(* IEC 61131-3 sources: s7-to-codesys/src/POUs/Lang/Converted/FB_PumpInterlockLad, 2 files *)

(* ---- FB_PumpInterlockLad.decl.st ---- *)
// Назначение: Блокировки насоса по уровню и давлению (LAD)
//             Блокировки насоса II подъёма по уровню в РЧВ и давлению в коллекторе (LAD).
//             1. xLowLevel := iLevel_cm < iLevelMin_cm.  2. xHighPress := iPressure_kPa > iPressureMax_kPa.
//             3. Если xLowLevel OR xHighPress — установить xAlarmLatch (S).
//             4. Если xAck AND NOT xLowLevel AND NOT xHighPress — сбросить xAlarmLatch (R).
//             5. Обслуживание: при xMaint прыжок вперёд к метке NoAuto (сети 6-7 не выполняются).
//             6. xPumpOn := xAutoReq AND NOT xAlarmLatch.
//             7. По фронту xPumpOn (P_TRIG, бит xRunEdge): iRunCount := iRunCount + 1 (ADD Int); xCountOk := ENO
//             сложения
//             (ENO = 0 при переполнении Int: 32767 + 1).
// Автор:      WTP2 (исходный блок S7); перевод в ST — s7conv 0.1.0
// Версия:     0.1 (исходный блок S7)
// Документ:   docs/CONVERSION_REPORT.md, docs/MAPPING.md
// Источник:   samples/lang/FB_PumpInterlockLad.xml, LAD, SW.Blocks.FB "FB_PumpInterlockLad", пространство имён
//             Interface/v5, FAMILY Drives
// Сгенерировано s7conv: пометки MIGRATION-CHECK и MIGRATION-TODO требуют ручного разбора.
FUNCTION_BLOCK FB_PumpInterlockLad
VAR_INPUT
    xAutoReq : BOOL;  // Запрос автоматики на работу
    iLevel_cm : INT;  // Уровень в РЧВ, см
    iLevelMin_cm : INT := 50;  // Минимальный уровень, см
    iPressure_kPa : INT;  // Давление в коллекторе, кПа
    iPressureMax_kPa : INT := 600;  // Максимальное давление, кПа
    xAck : BOOL;  // Квитирование аварии
    xMaint : BOOL;  // Режим обслуживания
END_VAR
VAR_OUTPUT
    xPumpOn : BOOL;  // Команда насосу
    xLowLevel : BOOL;  // Низкий уровень
    xHighPress : BOOL;  // Высокое давление
    xAlarm : BOOL;  // Авария (защёлка)
    iRunCount : INT;  // Число включений
    xCountOk : BOOL;  // ENO сложения: нет переполнения
    iSetpoint_pct : INT;  // Уставка производительности, %
    xChainOk : BOOL;  // ENO цепочки вызовов
    xRunMem : BOOL;  // Копия бита памяти фронта
END_VAR
VAR
    xAlarmLatch : BOOL;  // Защёлка аварии
    xRunEdge : BOOL;  // Бит памяти фронта xPumpOn
    iStage1 : INT;  // Уставка после первого ограничения
    iStage2 : INT;  // Уставка после второго ограничения
END_VAR
VAR_TEMP
    xNet5_1 : BOOL;  // сеть 5: условие прыжка к NoAuto (UId 21)
    xNet7_1 : BOOL;  // сеть 7: PBox (UId 21)
    xNet7_2 : BOOL;  // сеть 7: ENO Add (UId 25)
END_VAR

(* ---- FB_PumpInterlockLad.impl.st ---- *)
// Сеть 1: Низкий уровень в РЧВ
xLowLevel := iLevel_cm < iLevelMin_cm;
// Сеть 2: Высокое давление в коллекторе
xHighPress := iPressure_kPa > iPressureMax_kPa;
// Сеть 3: Защёлка аварии: установка
IF xLowLevel OR xHighPress THEN
    xAlarmLatch := TRUE;
END_IF
// Сеть 4: Защёлка аварии: квитирование
IF xAck AND NOT xLowLevel AND NOT xHighPress THEN
    xAlarmLatch := FALSE;
END_IF
// Сеть 5: Обслуживание: прыжок к NoAuto
// MIGRATION-CHECK: элемент «Jump»: имя и пины в SimaticML не подтверждены открытым экспортом
//                  (docs/MAPPING_LADFBD.md, уровень L) (FB_PumpInterlockLad.xml, сеть 5, UId 21)
xNet5_1 := xMaint;
IF NOT xNet5_1 THEN
    // прыжок к NoAuto: сети 6–7 выполняются без прыжка
    // Сеть 6: Автоматический режим
    xPumpOn := xAutoReq AND NOT xAlarmLatch;
    // Сеть 7: Счётчик включений с ENO
    xNet7_1 := xPumpOn AND NOT xRunEdge;
    xRunEdge := xPumpOn;
    // MIGRATION-CHECK: ENO Add S7 = EN AND NOT переполнение: F_S7EnoAddInt из S7Compat (в CODESYS ENO = EN);
    //                  результат при переполнении записывается с переносом, как у S7-300 [M]
    //                  (FB_PumpInterlockLad.xml, сеть 7, UId 25)
    xNet7_2 := xNet7_1 AND F_S7EnoAddInt(iIn1 := iRunCount, iIn2 := 1);
    IF xNet7_1 THEN
        iRunCount := iRunCount + 1;
    END_IF
    xCountOk := xNet7_2;
END_IF
// Сеть 8: Метка NoAuto: обслуживание выключает насос
IF xMaint THEN
    xPumpOn := FALSE;
END_IF
// Сеть 9: Уставка: три вызова FC_ClampPctLad через EN/ENO
// MIGRATION-CHECK: элемент «Call»: имя и пины в SimaticML не подтверждены открытым экспортом
//                  (docs/MAPPING_LADFBD.md, уровень L) (FB_PumpInterlockLad.xml, сеть 9, UId 23)
IF xPumpOn THEN
    iStage1 := FC_ClampPctLad(iIn := iLevel_cm, iMin := 0, iMax := 100);
END_IF
// MIGRATION-CHECK: элемент «Call»: имя и пины в SimaticML не подтверждены открытым экспортом
//                  (docs/MAPPING_LADFBD.md, уровень L) (FB_PumpInterlockLad.xml, сеть 9, UId 28)
IF xPumpOn THEN
    iStage2 := FC_ClampPctLad(iIn := iStage1, iMin := 10, iMax := 90);
END_IF
// MIGRATION-CHECK: элемент «Call»: имя и пины в SimaticML не подтверждены открытым экспортом
//                  (docs/MAPPING_LADFBD.md, уровень L) (FB_PumpInterlockLad.xml, сеть 9, UId 33)
IF xPumpOn THEN
    iSetpoint_pct := FC_ClampPctLad(iIn := iStage2, iMin := 20, iMax := 80);
END_IF
xChainOk := xPumpOn;
// Сеть 10: Насос выключен: уставка 0
IF NOT xPumpOn THEN
    iSetpoint_pct := 0;
END_IF
// Сеть 11: Авария
xAlarm := xAlarmLatch;
// Сеть 12: Бит памяти фронта в другой сети
xRunMem := xRunEdge;
